TYPE "DT_ALM_SYSTEM_WATERWAY"
VERSION : 0.1
   STRUCT
      MIV_LS_ERR { S7_SetPoint := 'False'} : "DT_ALM_SOLO" := (96, FALSE, TRUE, TRUE, (), (), 0, 3, 3, (), (), (), (), (), T#500MS);
      MIV_OPENING_TOO_LONG { S7_SetPoint := 'False'} : "DT_ALM_SOLO" := (97, FALSE, TRUE, TRUE, (), (), 0, 3, 3, (), (), (), (), (), T#3M);
      MIV_CLOSING_TOO_LONG { S7_SetPoint := 'False'} : "DT_ALM_SOLO" := (98, FALSE, TRUE, TRUE, (), (), 0, 3, 3, (), (), (), (), (), T#3M);
      MIV_SELFCLOSURE { S7_SetPoint := 'False'} : "DT_ALM_SOLO" := (99, FALSE, TRUE, TRUE, (), (), 0, 3, 3, (), (), (), (), (), T#10S);
      MIV_OPENING_TOO_SHORT { S7_SetPoint := 'False'} : "DT_ALM_SOLO" := (100, FALSE, FALSE, FALSE, (), (), 0, 0, 0, (), (), (), (), (), T#500MS);
      MIV_CLOSING_TOO_SHORT { S7_SetPoint := 'False'} : "DT_ALM_SOLO" := (101, FALSE, FALSE, FALSE, (), (), 0, 0, 0, (), (), (), (), (), T#500MS);
      MIV_SAFETY_PIN { S7_SetPoint := 'False'} : "DT_ALM_SOLO" := (102, FALSE, FALSE, FALSE, (), (), 0, 0, 0, (), (), (), (), (), T#500MS);
      BYP_LS_ERR { S7_SetPoint := 'False'} : "DT_ALM_SOLO" := (103, FALSE, TRUE, TRUE, (), (), 0, 3, 0, (), (), (), (), (), T#500MS);
      BYP_OPENING_TOO_LONG { S7_SetPoint := 'False'} : "DT_ALM_SOLO" := (104, FALSE, TRUE, TRUE, (), (), 0, 3, 0, (), (), (), (), (), T#1M);
      BYP_CLOSING_TOO_LONG { S7_SetPoint := 'False'} : "DT_ALM_SOLO" := (105, FALSE, TRUE, TRUE, (), (), 0, 3, 0, (), (), (), (), (), T#1M);
      BYP_MCB_OFF { S7_SetPoint := 'False'} : "DT_ALM_SOLO" := (106, FALSE, TRUE, TRUE, (), (), 1, 0, 1, (), (), (), (), (), T#500MS);
      BYP_CONT_OP_ERR { S7_SetPoint := 'False'} : "DT_ALM_SOLO" := (107, FALSE, TRUE, TRUE, (), (), 1, 0, 2, (), (), (), (), (), T#2S);
      BYP_CONT_CL_ERR { S7_SetPoint := 'False'} : "DT_ALM_SOLO" := (108, FALSE, TRUE, TRUE, (), (), 1, 0, 2, (), (), (), (), (), T#2S);
      BYP_TORQUE_OP { S7_SetPoint := 'False'} : "DT_ALM_SOLO" := (109, FALSE, TRUE, TRUE, (), (), 1, 0, 3, (), (), (), (), (), T#500MS);
      BYP_TORQUE_CL { S7_SetPoint := 'False'} : "DT_ALM_SOLO" := (110, FALSE, FALSE, FALSE, (), (), 0, 0, 0, (), (), (), (), (), T#500MS);
      BYP_TH_OVERLOAD { S7_SetPoint := 'False'} : "DT_ALM_SOLO" := (111, FALSE, FALSE, FALSE, (), (), 0, 0, 0, (), (), (), (), (), T#500MS);
      BYP_HEAT_MCB_OFF { S7_SetPoint := 'False'} : "DT_ALM_SOLO" := (112, FALSE, FALSE, FALSE, (), (), 0, 0, 0, (), (), (), (), (), T#500MS);
      PENSTOCK_ERR { S7_SetPoint := 'False'} : "DT_ALM_SOLO" := (113, FALSE, TRUE, TRUE, (), (), 0, 2, 2, (), (), (), (), (), T#3S);
      PENSTOCK_PRESSURE_LL { S7_SetPoint := 'False'} : "DT_ALM_SOLO" := (114, FALSE, TRUE, TRUE, (), (), 0, 2, 3, (), (), (), (), (), T#5S);
      PENSTOCK_PRESSURE_L { S7_SetPoint := 'False'} : "DT_ALM_SOLO" := (115, FALSE, TRUE, TRUE, (), (), 0, 2, 1, (), (), (), (), (), T#5S);
      TURBINE_ERR { S7_SetPoint := 'False'} : "DT_ALM_SOLO" := (116, FALSE, TRUE, TRUE, (), (), 0, 2, 2, (), (), (), (), (), T#3S);
      TURBINE_PRESSURE_LL { S7_SetPoint := 'False'} : "DT_ALM_SOLO" := (117, FALSE, TRUE, TRUE, (), (), 0, 2, 3, (), (), (), (), (), T#5S);
      TURBINE_PRESSURE_L { S7_SetPoint := 'False'} : "DT_ALM_SOLO" := (118, FALSE, TRUE, TRUE, (), (), 0, 2, 1, (), (), (), (), (), T#5S);
      DIFF_PRESSURE { S7_SetPoint := 'False'} : "DT_ALM_SOLO" := (119, FALSE, FALSE, FALSE, (), (), 0, 0, 0, (), (), (), (), (), T#500MS);
      BYP_CONT_ERR { S7_SetPoint := 'False'} : "DT_ALM_SOLO" := (120, FALSE, FALSE, FALSE, (), (), 0, 0, 0, (), (), (), (), (), T#500MS);
      MIV_MCB_OFF { S7_SetPoint := 'False'} : "DT_ALM_SOLO" := (121, FALSE, FALSE, TRUE, (), (), 1, 0, 3, (), (), (), (), (), T#500MS);
      MIV_CONT_ERR { S7_SetPoint := 'False'} : "DT_ALM_SOLO" := (122, FALSE, FALSE, TRUE, (), (), 1, 0, 3, (), (), (), (), (), T#2S);
      MIV_HEAT_MCB_OFF { S7_SetPoint := 'False'} : "DT_ALM_SOLO" := (123, FALSE, FALSE, TRUE, (), (), 1, 0, 3, (), (), (), (), (), T#500MS);
      MIV_TORQUE_OP { S7_SetPoint := 'False'} : "DT_ALM_SOLO" := (124, FALSE, FALSE, TRUE, (), (), 1, 3, 3, (), (), (), (), (), T#500MS);
      MIV_TORQUE_CL { S7_SetPoint := 'False'} : "DT_ALM_SOLO" := (125, FALSE, FALSE, TRUE, (), (), 1, 3, 3, (), (), (), (), (), T#500MS);
      MIV_TH_OVERLOAD { S7_SetPoint := 'False'} : "DT_ALM_SOLO" := (126, FALSE, FALSE, TRUE, (), (), 1, 3, 3, (), (), (), (), (), T#500MS);
      SPARE_127 { S7_SetPoint := 'False'} : "DT_ALM_SOLO" := (127, FALSE, FALSE, FALSE, (), (), 0, 0, 0, (), (), (), (), (), T#500MS);
   END_STRUCT;

END_TYPE

